Fanuc KAREL source: kb00007.KL

PROGRAM KB00007
%STACKSIZE=65535
%PRIORITY=65535
%NOLOCKGROUP
VAR
P1 : POSITION
RESULT : VECTOR
BEGIN
RESULT=APPROACH(P1)
END KB00007
